SUBAPPLICATION TestSubApp (* Subapplication with a basic FB *)
  (* Standard: 61499-1; Description: Copyright (c) 2026 Martin Erich Jobst This program and the accompanying materials are made available under the terms of the Eclipse Public License 2.0 which is available at https://www.eclipse.org/legal/epl-2.0/ SPDX-License-Identifier: EPL-2.0 *)
  (* Version 1.0, 2026-10-23, Martin Jobst *)
  {SET_ATTRIBUTE(IntegerAttribute, 17)}
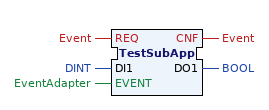
  EVENT_INPUT
    REQ; (* Request *)
  END_EVENT
  EVENT_OUTPUT
    CNF; (* Confirmation *)
  END_EVENT
  VAR_INPUT
    DI1 : DINT := DINT#5;
  END_VAR
  VAR_OUTPUT
    DO1 : BOOL;
  END_VAR
  SOCKETS
    EVENT : EventAdapter; (* Event/data adapter *)
  END_SOCKETS
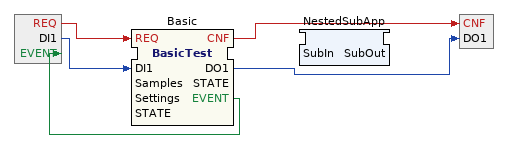
  (* Subapplication network comment *)
  FBS
    Basic : fixture::basic::BasicTest;
  END_FBS
  SUBAPPLICATION NestedSubApp
    {SET_ATTRIBUTE(IntegerAttribute, 16)}
    {SET_ATTRIBUTE(locked, true)}
    VAR_INPUT
      SubIn : DINT;
    END_VAR
    VAR_OUTPUT
      SubOut : BOOL;
    END_VAR
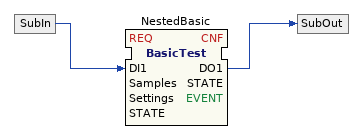
    FBS
      NestedBasic : fixture::basic::BasicTest;
    END_FBS
    DATA_CONNECTIONS
      SubIn TO NestedBasic.DI1;
      NestedBasic.DO1 TO SubOut;
    END_CONNECTIONS
  END_SUBAPPLICATION
  EVENT_CONNECTIONS
    REQ TO Basic.REQ;
    Basic.CNF TO CNF;
  END_CONNECTIONS
  DATA_CONNECTIONS
    DI1 TO Basic.DI1;
    Basic.DO1 TO DO1;
  END_CONNECTIONS
  ADAPTER_CONNECTIONS
    Basic.EVENT TO EVENT;
  END_CONNECTIONS
END_SUBAPPLICATION
